GLOBALCONSTANTS SubStrings (* Global constants *)
  (* Standard: 61499-1 *)
  (* Version 1.0, 2026-11-06, Franz Höpfinger, Meisterschulen am Ostbahnhof *)
  PACKAGE Meins::Servo_AI3_Calibrate_2P_OPC;
  VAR_GLOBAL CONSTANT
    SAI3_RAW_WRITE : WSTRING := "opc_ua[WRITE;/Objects/ServoAI3/RAW,1:s=SAI3_RAW]"; (* Rohwert AI3 0-4095 *)
    SAI3_CAL_WRITE : WSTRING := "opc_ua[WRITE;/Objects/ServoAI3/CAL,1:s=SAI3_CAL]"; (* kalibrierter Wert AI3 = Sollwinkel *)
    SAI3_CO_METHOD : WSTRING := "opc_ua[CREATE_METHOD;/Objects/ServoAI3/COMethod,1:s=SAI3_CO_METHOD]"; (* Trigger CO (Nullpunkt) *)
    SAI3_CS_METHOD : WSTRING := "opc_ua[CREATE_METHOD;/Objects/ServoAI3/CSMethod,1:s=SAI3_CS_METHOD]"; (* Trigger CS (Spanne) *)
    SAI3_ZERO_READ : WSTRING := "opc_ua[READ;/Objects/ServoAI3/ZEROREFExt,1:s=SAI3_ZEROREF_EXT]"; (* ZERO_REF vom Dashboard *)
    SAI3_ZERO_WRITE : WSTRING := "opc_ua[WRITE;/Objects/ServoAI3/ZEROREF,1:s=SAI3_ZEROREF]"; (* ZERO_REF Echo *)
    SAI3_SPAN_READ : WSTRING := "opc_ua[READ;/Objects/ServoAI3/SPANREFExt,1:s=SAI3_SPANREF_EXT]"; (* SPAN_REF vom Dashboard *)
    SAI3_SPAN_WRITE : WSTRING := "opc_ua[WRITE;/Objects/ServoAI3/SPANREF,1:s=SAI3_SPANREF]"; (* SPAN_REF Echo *)
    SAI3_ZERO_RAW_WRITE : WSTRING := "opc_ua[WRITE;/Objects/ServoAI3/ZERORAW,1:s=SAI3_ZERO_RAW]"; (* Rohwert am ZERO-Punkt *)
    SAI3_SPAN_RAW_WRITE : WSTRING := "opc_ua[WRITE;/Objects/ServoAI3/SPANRAW,1:s=SAI3_SPAN_RAW]"; (* Rohwert am SPAN-Punkt *)
    SAI3_ANGLE : WSTRING := "opc_ua[WRITE;/Objects/ServoAI3/ANGLE,1:s=SAI3_ANGLE]"; (* angewendeter Winkel Q2 (Echo) *)
  END_VAR
END_GLOBALCONSTANTS
